Fanuc KAREL source: ka00195.KL

PROGRAM KA00195
%STACKSIZE=65535
%PRIORITY=65535
%NOLOCKGROUP
VAR
SRC : ARRAY[4] OF SHORT
DST : ARRAY[4] OF SHORT
BEGIN
-- UNRESOLVED_PC line 7 opcodes [22 22 1E] marker_code=0
END KA00195
